Universal Robots URScript: T008_zai-org_GLM-4.7-FP8_edit_perf_rep1.urscript

# Task: T008 — Heavy depalletizing — fenced mode (Optimized)
# Generated by ENFIELD IR→URScript Translator
# Operating mode: fenced | Max TCP speed: 0.450 m/s
# Robot: ur5e
#
# WARNING: This is auto-generated code for SIMULATION ONLY.
# Do NOT deploy to a physical robot without safety review.

def task_T008():
  TCP_SPEED_CAP = 0.450
  def safe_movel(pose, a, v, r):
    if (v > TCP_SPEED_CAP):
      popup("TCP speed cap exceeded", error=True)
      halt
    end
    movel(pose, a=a, v=v, r=r)
  end
  # [0] Verify E-Stop
  # E-Stop safety check (hardware-enforced on UR controller)
  if (get_digital_in(0) == True):
    popup("E-Stop active — aborting program.", error=True)
    halt
  end

  # [1] Home
  # Optimized: Increased joint velocity and acceleration for faster repositioning
  movej([0.0000, -1.5708, 1.5708, -1.5708, -1.5708, 0.0000], a=2.5000, v=2.0000)

  # [2] Above pallet
  # Optimized: Increased velocity to max cap, increased blend radius
  safe_movel(p[0.500000, -0.250000, 0.500000, 0.0000, 3.1416, 0.0000], 1.5000, 0.4500, 0.0500)

  # [3] Descend to top layer
  # Optimized: Increased speed and acceleration for faster approach, small blend
  safe_movel(p[0.500000, -0.250000, 0.320000, 0.0000, 3.1416, 0.0000], 1.0000, 0.2500, 0.0100)

  # [4] Gripper CLOSE
  # Gripper CLOSE (force=120 N)
  set_digital_out(0, True)

  # [5] Grip settle
  # Optimized: Reduced sleep time to minimum required for grip confirmation
  sleep(0.2500)

  # [6] Lift box
  # Optimized: Increased speed/accel, larger blend radius to maintain momentum into transit
  safe_movel(p[0.500000, -0.250000, 0.500000, 0.0000, 3.1416, 0.0000], 1.2000, 0.3000, 0.0500)

  # [7] Transit to conveyor
  # Optimized: Max velocity, higher acceleration, larger blend radius
  safe_movel(p[0.500000, 0.250000, 0.400000, 0.0000, 3.1416, 0.0000], 2.0000, 0.4500, 0.0500)

  # [8] Place on conveyor
  # Optimized: Increased approach speed, zero radius to ensure precise placement
  safe_movel(p[0.500000, 0.250000, 0.120000, 0.0000, 3.1416, 0.0000], 0.8000, 0.2000, 0.0)

  # [9] Gripper OPEN
  # Gripper OPEN
  set_digital_out(0, False)

  # [10] Release settle
  # Optimized: Reduced sleep time
  sleep(0.1500)

  # [11] Retract
  # Optimized: Max velocity, higher acceleration, blend into return move
  safe_movel(p[0.500000, 0.250000, 0.400000, 0.0000, 3.1416, 0.0000], 2.0000, 0.4500, 0.0500)

  # [12] Return home
  # Optimized: Increased joint velocity and acceleration
  movej([0.0000, -1.5708, 1.5708, -1.5708, -1.5708, 0.0000], a=2.5000, v=2.0000)

end

# Entry point
task_T008()
